(* Logix 5000 project; controller TFF vendor 1 type 14 code 107 rev 33.11; software revision 33.04; part 25 of 38 *)
(* tags used below, declared in another part *)
   Address : DINT;   // Temp Address
   Address2 : DINT;   // Temp Address
   Index : DINT;   // Index
   PCV001_PID_Settings : INT;
   TIME : DINT[2];
   AnalogOutput : AnalogOutput[25];   // Analog Output Array
   AnalogPoint : AnalogInput[50];   // Analog Input Array
   ControlLoop : ControlLoop[20];   // Control Loop Array
   ControlLoop_FeedPump : ALIAS FOR ControlLoop[1];
   ControlLoop_PCV101 : ALIAS FOR ControlLoop[3];
   ControlLoop_PCV101_5ms : ALIAS FOR ControlLoop[4];
   ControlLoop_PCV101_CV : REAL;   // Control Value
   ControlLoop_PCV101_RAMP_OUT : REAL;   // Ramp Output
   ControlLoop_PCV201 : ALIAS FOR ControlLoop[5];
   ControlLoop_PCV201_5ms : ALIAS FOR ControlLoop[6];
   ControlLoop_PCV201_RAMP_OUT : REAL;   // Ramp Output
   PCV101 : ALIAS FOR AnalogPoint[3];
   PCV101_Control : PCV_Control;   // PCV101 Control UDT
   PCV201_Control : PCV_Control;   // PCV201 Control UDT
   PumpRunStatus : DINT;   // Pumps Run Status (1 = At least one pump running , 0 = no pump running)
   SysControl : SysControl;   // General system status and command
(* Process, continued *)

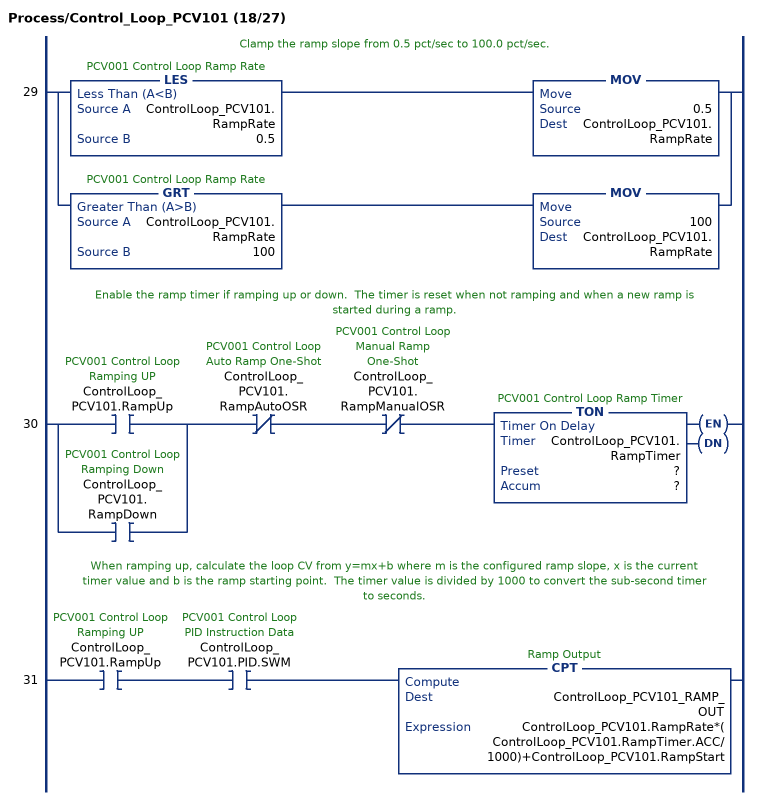
   [picture p215: Process/Control_Loop_PCV101 rungs 29-31]
   // Clamp the ramp slope from 0.5 pct/sec to 100.0 pct/sec.
   29: [LES(ControlLoop_PCV101.RampRate,0.5) MOV(0.5,ControlLoop_PCV101.RampRate) ,GRT(ControlLoop_PCV101.RampRate,100) MOV(100,ControlLoop_PCV101.RampRate) ];
   // Enable the ramp timer if ramping up or down.  The timer is reset when not ramping and when a new ramp is started during a ramp.
   30: [XIC(ControlLoop_PCV101.RampUp) ,XIC(ControlLoop_PCV101.RampDown) ]XIO(ControlLoop_PCV101.RampAutoOSR)XIO(ControlLoop_PCV101.RampManualOSR)TON(ControlLoop_PCV101.RampTimer,?,?);
   // When ramping up, calculate the loop CV from y=mx+b where m is the configured ramp slope, x is the current timer value and b is the ramp starting point.  The timer value is divided by 1000 to convert the sub-second timer to seconds.
   31: XIC(ControlLoop_PCV101.RampUp)XIC(ControlLoop_PCV101.PID.SWM)CPT(ControlLoop_PCV101_RAMP_OUT,ControlLoop_PCV101.RampRate*(ControlLoop_PCV101.RampTimer.ACC/1000)+ControlLoop_PCV101.RampStart);
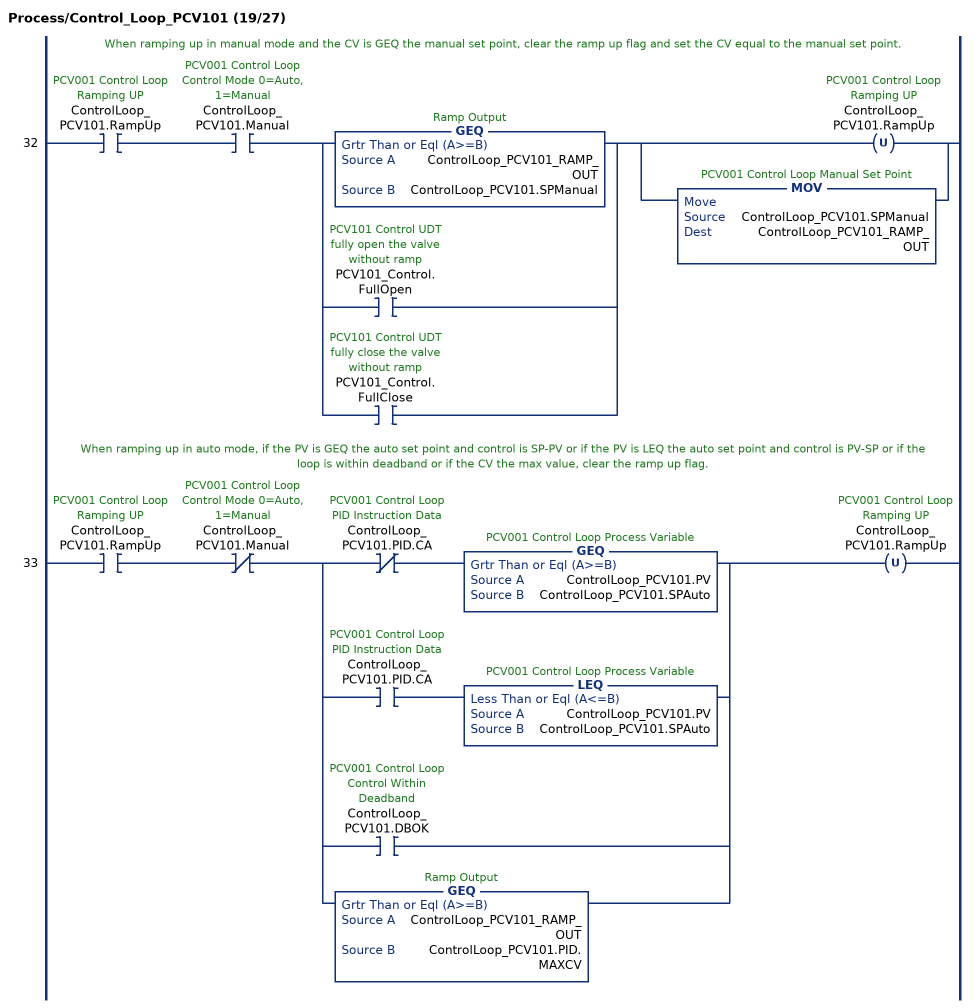
   // When ramping up in manual mode and the CV is GEQ the manual set point, clear the ramp up flag and set the CV equal to the manual set point.
   32: XIC(ControlLoop_PCV101.RampUp)XIC(ControlLoop_PCV101.Manual)[GEQ(ControlLoop_PCV101_RAMP_OUT,ControlLoop_PCV101.SPManual) ,XIC(PCV101_Control.FullOpen) ,XIC(PCV101_Control.FullClose) ][OTU(ControlLoop_PCV101.RampUp) ,MOV(ControlLoop_PCV101.SPManual,ControlLoop_PCV101_RAMP_OUT) ];
   // When ramping up in auto mode, if the PV is GEQ the auto set point and control is SP-PV or if the PV is LEQ the auto set point and control is PV-SP or if the loop is within deadband or if the CV the max value, clear the ramp up flag.
   33: XIC(ControlLoop_PCV101.RampUp)XIO(ControlLoop_PCV101.Manual)[XIO(ControlLoop_PCV101.PID.CA) GEQ(ControlLoop_PCV101.PV,ControlLoop_PCV101.SPAuto) ,XIC(ControlLoop_PCV101.PID.CA) LEQ(ControlLoop_PCV101.PV,ControlLoop_PCV101.SPAuto) ,XIC(ControlLoop_PCV101.DBOK) ,GEQ(ControlLoop_PCV101_RAMP_OUT,ControlLoop_PCV101.PID.MAXCV) ]OTU(ControlLoop_PCV101.RampUp);
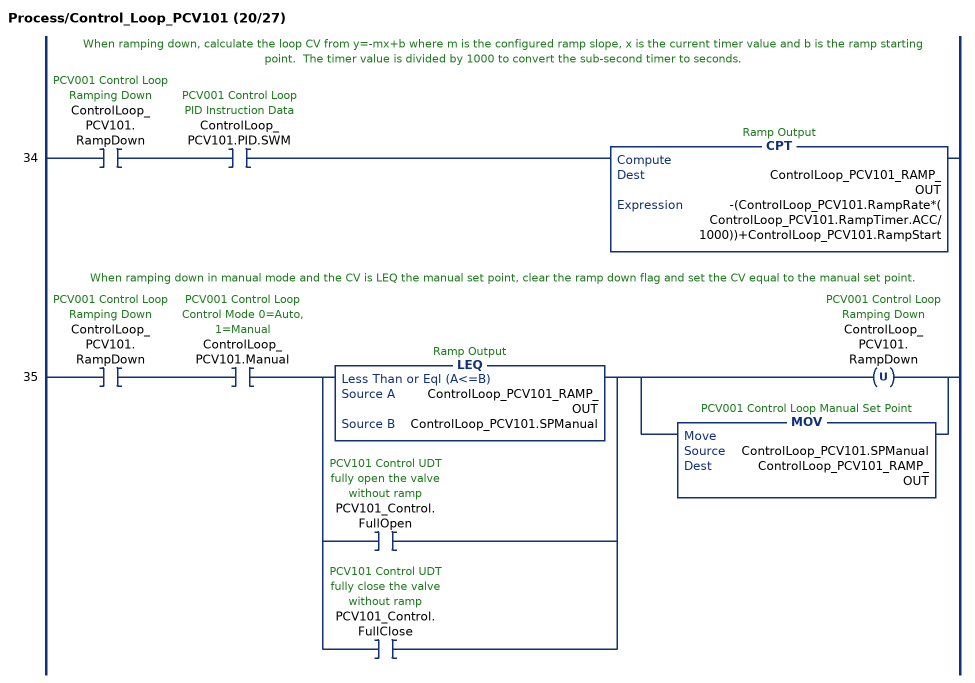
   // When ramping down, calculate the loop CV from y=-mx+b where m is the configured ramp slope, x is the current timer value and b is the ramp starting point.  The timer value is divided by 1000 to convert the sub-second timer to seconds.
   34: XIC(ControlLoop_PCV101.RampDown)XIC(ControlLoop_PCV101.PID.SWM)CPT(ControlLoop_PCV101_RAMP_OUT,-(ControlLoop_PCV101.RampRate*(ControlLoop_PCV101.RampTimer.ACC/1000))+ControlLoop_PCV101.RampStart);
   // When ramping down in manual mode and the CV is LEQ the manual set point, clear the ramp down flag and set the CV equal to the manual set point.
   35: XIC(ControlLoop_PCV101.RampDown)XIC(ControlLoop_PCV101.Manual)[LEQ(ControlLoop_PCV101_RAMP_OUT,ControlLoop_PCV101.SPManual) ,XIC(PCV101_Control.FullOpen) ,XIC(PCV101_Control.FullClose) ][OTU(ControlLoop_PCV101.RampDown) ,MOV(ControlLoop_PCV101.SPManual,ControlLoop_PCV101_RAMP_OUT) ];
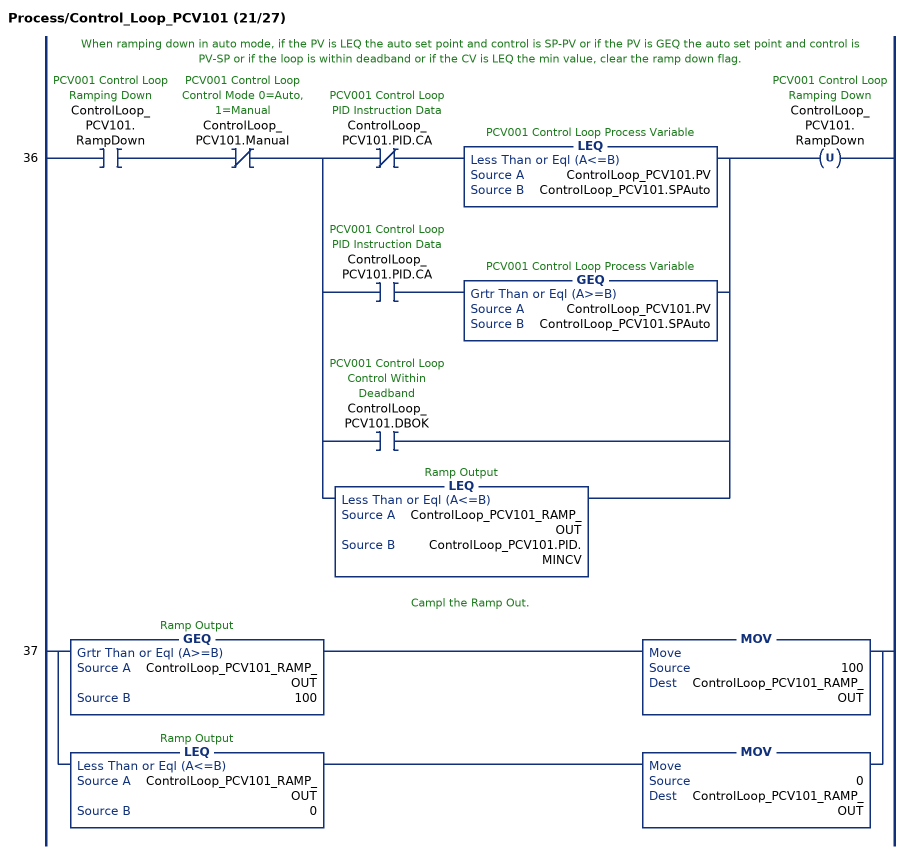
   // When ramping down in auto mode, if the PV is LEQ the auto set point and control is SP-PV or if the PV is GEQ the auto set point and control is PV-SP or if the loop is within deadband or if the CV is LEQ the min value, clear the ramp down flag.
   36: XIC(ControlLoop_PCV101.RampDown)XIO(ControlLoop_PCV101.Manual)[XIO(ControlLoop_PCV101.PID.CA) LEQ(ControlLoop_PCV101.PV,ControlLoop_PCV101.SPAuto) ,XIC(ControlLoop_PCV101.PID.CA) GEQ(ControlLoop_PCV101.PV,ControlLoop_PCV101.SPAuto) ,XIC(ControlLoop_PCV101.DBOK) ,LEQ(ControlLoop_PCV101_RAMP_OUT,ControlLoop_PCV101.PID.MINCV) ]OTU(ControlLoop_PCV101.RampDown);
   // Campl the Ramp Out.
   37: [GEQ(ControlLoop_PCV101_RAMP_OUT,100) MOV(100,ControlLoop_PCV101_RAMP_OUT) ,LEQ(ControlLoop_PCV101_RAMP_OUT,0) MOV(0,ControlLoop_PCV101_RAMP_OUT) ];
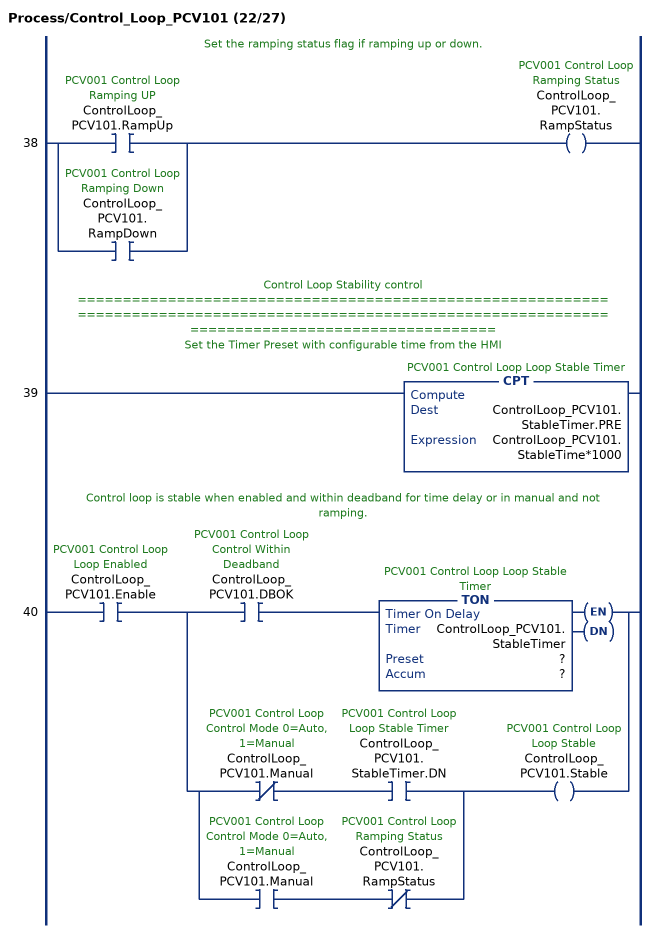
   // Set the ramping status flag if ramping up or down.
   38: [XIC(ControlLoop_PCV101.RampUp) ,XIC(ControlLoop_PCV101.RampDown) ]OTE(ControlLoop_PCV101.RampStatus);
   // Control Loop Stability control
   // ========================================================================================================================================================
   // Set the Timer Preset with configurable time from the HMI
   39: CPT(ControlLoop_PCV101.StableTimer.PRE,ControlLoop_PCV101.StableTime*1000);
   // Control loop is stable when enabled and within deadband for time delay or in manual and not ramping.
   40: XIC(ControlLoop_PCV101.Enable)[XIC(ControlLoop_PCV101.DBOK) TON(ControlLoop_PCV101.StableTimer,?,?) ,[XIO(ControlLoop_PCV101.Manual) XIC(ControlLoop_PCV101.StableTimer.DN) ,XIC(ControlLoop_PCV101.Manual) XIO(ControlLoop_PCV101.RampStatus) ] OTE(ControlLoop_PCV101.Stable) ];
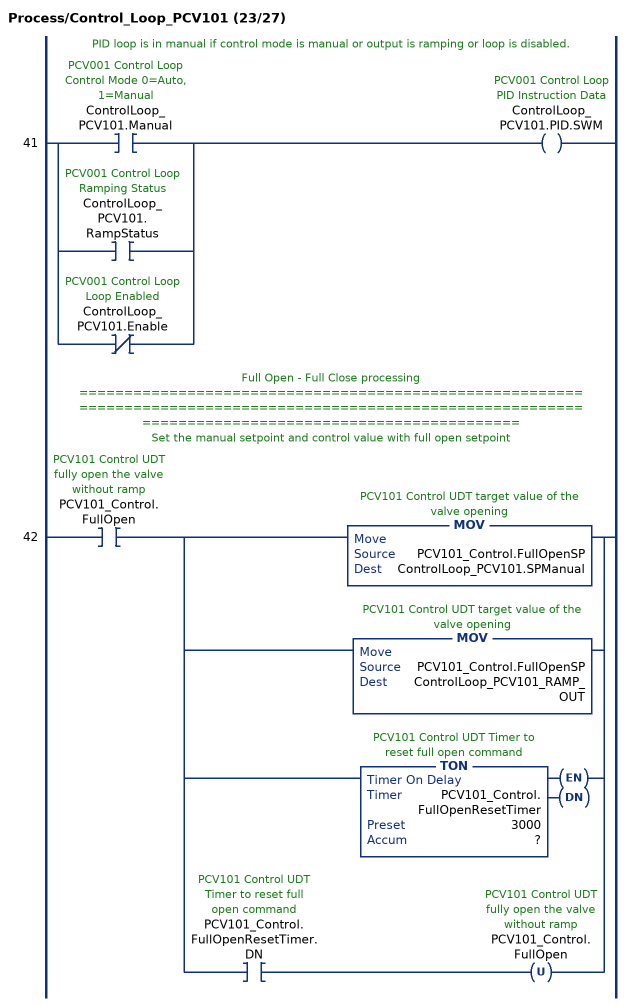
   // PID loop is in manual if control mode is manual or output is ramping or loop is disabled.
   41: [XIC(ControlLoop_PCV101.Manual) ,XIC(ControlLoop_PCV101.RampStatus) ,XIO(ControlLoop_PCV101.Enable) ]OTE(ControlLoop_PCV101.PID.SWM);
   // Full Open - Full Close processing
   // ==========================================================================================================================================================
   // Set the manual setpoint and control value with full open setpoint
   42: XIC(PCV101_Control.FullOpen)[MOV(PCV101_Control.FullOpenSP,ControlLoop_PCV101.SPManual) ,MOV(PCV101_Control.FullOpenSP,ControlLoop_PCV101_RAMP_OUT) ,TON(PCV101_Control.FullOpenResetTimer,?,?) ,XIC(PCV101_Control.FullOpenResetTimer.DN) OTU(PCV101_Control.FullOpen) ];
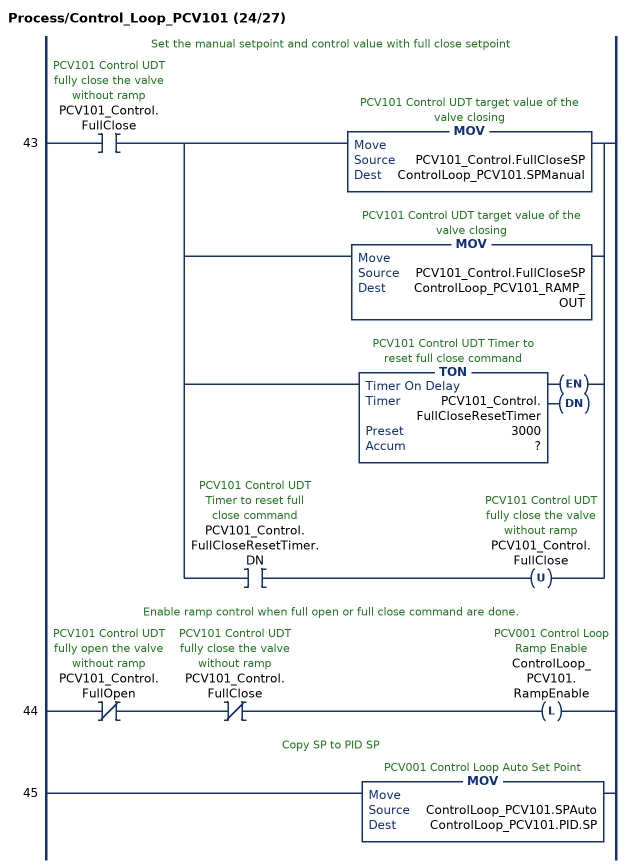
   // Set the manual setpoint and control value with full close setpoint
   43: XIC(PCV101_Control.FullClose)[MOV(PCV101_Control.FullCloseSP,ControlLoop_PCV101.SPManual) ,MOV(PCV101_Control.FullCloseSP,ControlLoop_PCV101_RAMP_OUT) ,TON(PCV101_Control.FullCloseResetTimer,?,?) ,XIC(PCV101_Control.FullCloseResetTimer.DN) OTU(PCV101_Control.FullClose) ];
   // Enable ramp control when full open or full close command are done.
   44: XIO(PCV101_Control.FullOpen)XIO(PCV101_Control.FullClose)OTL(ControlLoop_PCV101.RampEnable);
   // Copy SP to PID SP
   45: MOV(ControlLoop_PCV101.SPAuto,ControlLoop_PCV101.PID.SP);
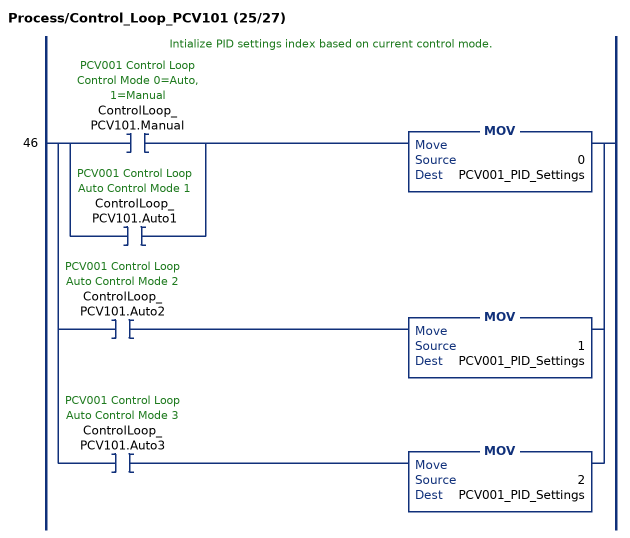
   // Intialize PID settings index based on current control mode.
   46: [[XIC(ControlLoop_PCV101.Manual) ,XIC(ControlLoop_PCV101.Auto1) ] MOV(0,PCV001_PID_Settings) ,XIC(ControlLoop_PCV101.Auto2) MOV(1,PCV001_PID_Settings) ,XIC(ControlLoop_PCV101.Auto3) MOV(2,PCV001_PID_Settings) ];
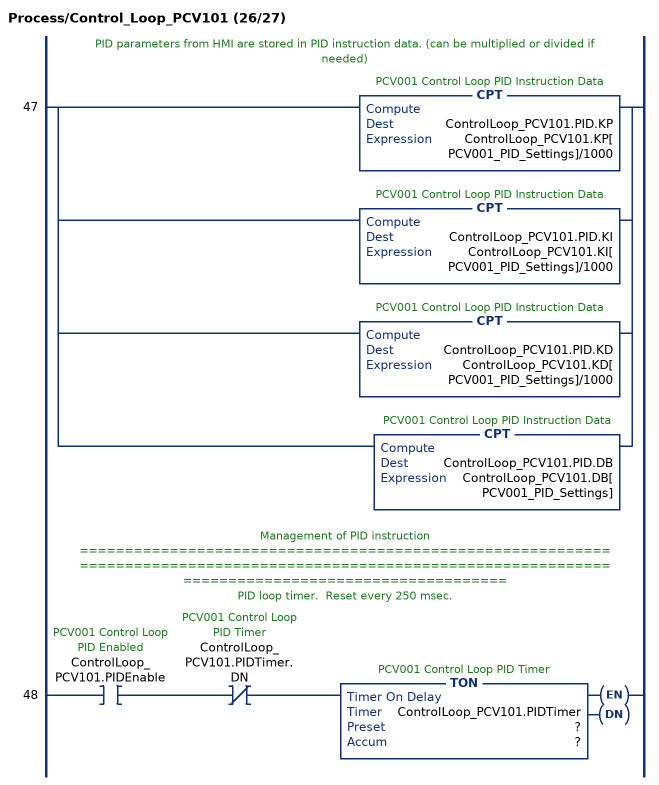
   // PID parameters from HMI are stored in PID instruction data. (can be multiplied or divided if needed)
   47: [CPT(ControlLoop_PCV101.PID.KP,ControlLoop_PCV101.KP[PCV001_PID_Settings]/1000) ,CPT(ControlLoop_PCV101.PID.KI,ControlLoop_PCV101.KI[PCV001_PID_Settings]/1000) ,CPT(ControlLoop_PCV101.PID.KD,ControlLoop_PCV101.KD[PCV001_PID_Settings]/1000) ,CPT(ControlLoop_PCV101.PID.DB,ControlLoop_PCV101.DB[PCV001_PID_Settings]) ];
   // Management of PID instruction
   // ==========================================================================================================================================================
   // PID loop timer.  Reset every 250 msec.
   48: XIC(ControlLoop_PCV101.PIDEnable)XIO(ControlLoop_PCV101.PIDTimer.DN)TON(ControlLoop_PCV101.PIDTimer,?,?);
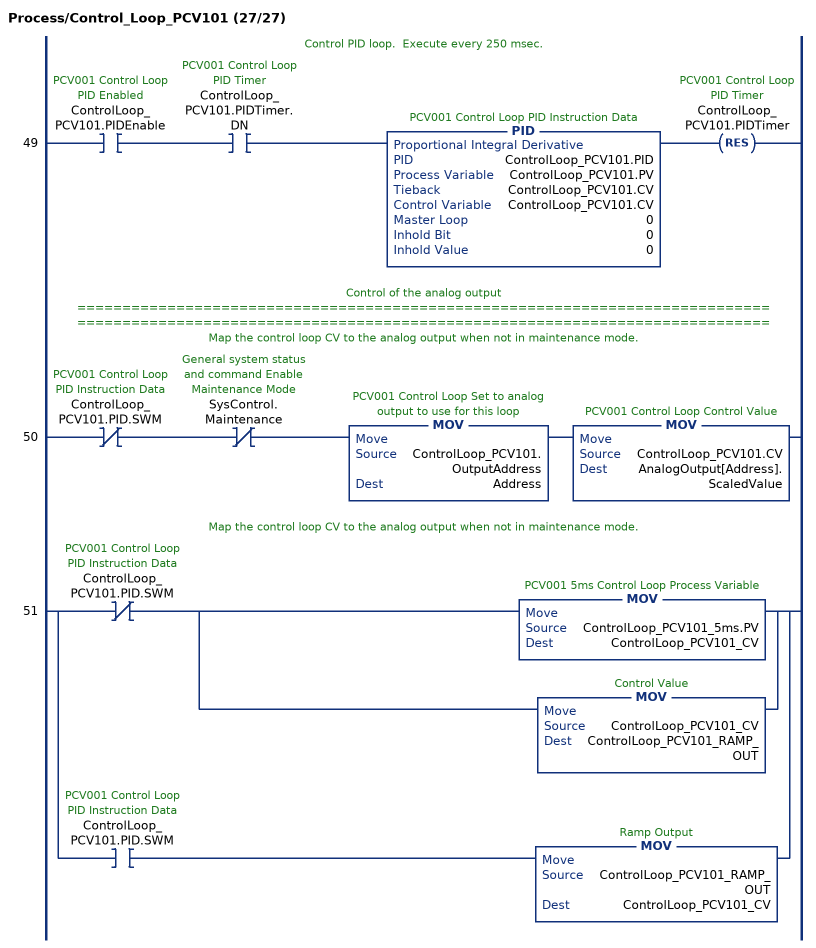
   // Control PID loop.  Execute every 250 msec.
   49: XIC(ControlLoop_PCV101.PIDEnable)XIC(ControlLoop_PCV101.PIDTimer.DN)PID(ControlLoop_PCV101.PID,ControlLoop_PCV101.PV,ControlLoop_PCV101.CV,ControlLoop_PCV101.CV,0,0,0)RES(ControlLoop_PCV101.PIDTimer);
   // Control of the analog output
   // ==========================================================================================================================================================
   // Map the control loop CV to the analog output when not in maintenance mode.
   50: XIO(ControlLoop_PCV101.PID.SWM)XIO(SysControl.Maintenance)MOV(ControlLoop_PCV101.OutputAddress,Address)MOV(ControlLoop_PCV101.CV,AnalogOutput[Address].ScaledValue);
   // Map the control loop CV to the analog output when not in maintenance mode.
   51: [XIO(ControlLoop_PCV101.PID.SWM) [MOV(ControlLoop_PCV101_5ms.PV,ControlLoop_PCV101_CV) ,MOV(ControlLoop_PCV101_CV,ControlLoop_PCV101_RAMP_OUT) ] ,XIC(ControlLoop_PCV101.PID.SWM) MOV(ControlLoop_PCV101_RAMP_OUT,ControlLoop_PCV101_CV) ];
END_ROUTINE

ROUTINE Control_Loop_PCV201   (* ladder *)
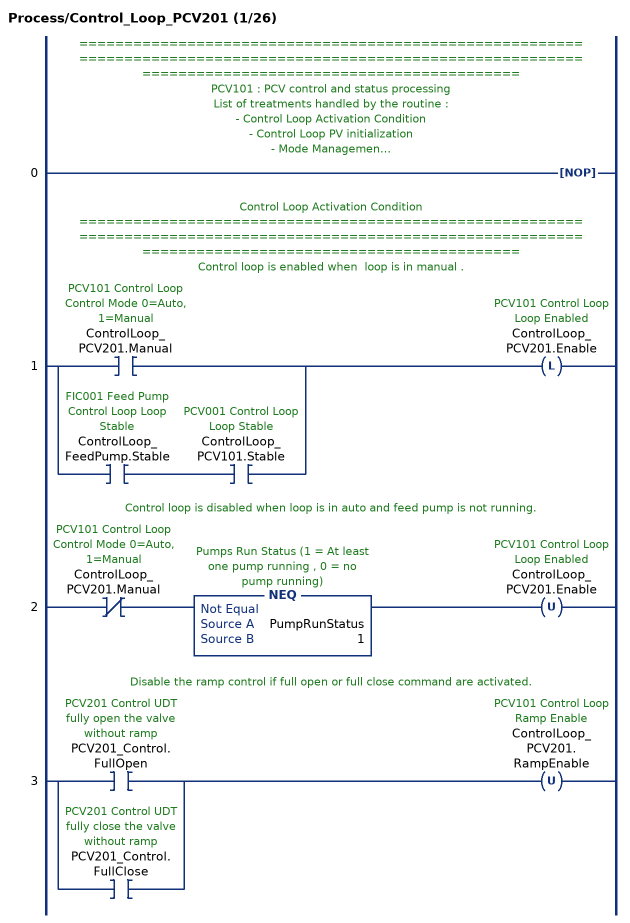
   // ==========================================================================================================================================================
   //                                                  PCV101 : PCV control and status processing
   //                                                     List of treatments handled by the routine :
   //                                                          - Control Loop Activation Condition
   //                                                  - Control Loop PV initialization
   //                                                - Mode Management
   //                                                        - Control Loop Setpoint management
   //                                                        - Control Loop deadband calculation
   //                                                          - Management of ramping control
   //                                                          - Control Loop Stability control
   //                                                          - Full Open - Full Close processing
   //                                                          - Management of PID instruction
   //                                                          - Control of the analog output
   //                                                     -----------------------------------------------------------------------------------------------------------------------------------------------------
   //                                                     History
   // 		2019-DEC-24 - Merck - Q. Spindler - Initial version for Candidate Release 1.00.00.00.a
   // 		2020-SEP-09 - Merck - Q. Spindler - Modifications for Candidate Release 1.00.00.00.d
   // 					- Add ControlLoop Enable and not manual condition for DBOK status
   // 		2021-APR-16 - Merck - Q. Spindler - Modifications for Candidate Release 1.00.00.00.e
   //                                        - Add Initialize address if no mode selected.
   // ==========================================================================================================================================================
   0: NOP();
   // Control Loop Activation Condition
   // ==========================================================================================================================================================
   // Control loop is enabled when  loop is in manual .
   1: [XIC(ControlLoop_PCV201.Manual) ,XIC(ControlLoop_FeedPump.Stable) XIC(ControlLoop_PCV101.Stable) ]OTL(ControlLoop_PCV201.Enable);
   // Control loop is disabled when loop is in auto and feed pump is not running.
   2: XIO(ControlLoop_PCV201.Manual)NEQ(PumpRunStatus,1)OTU(ControlLoop_PCV201.Enable);
   // Disable the ramp control if full open or full close command are activated.
   3: [XIC(PCV201_Control.FullOpen) ,XIC(PCV201_Control.FullClose) ]OTU(ControlLoop_PCV201.RampEnable);
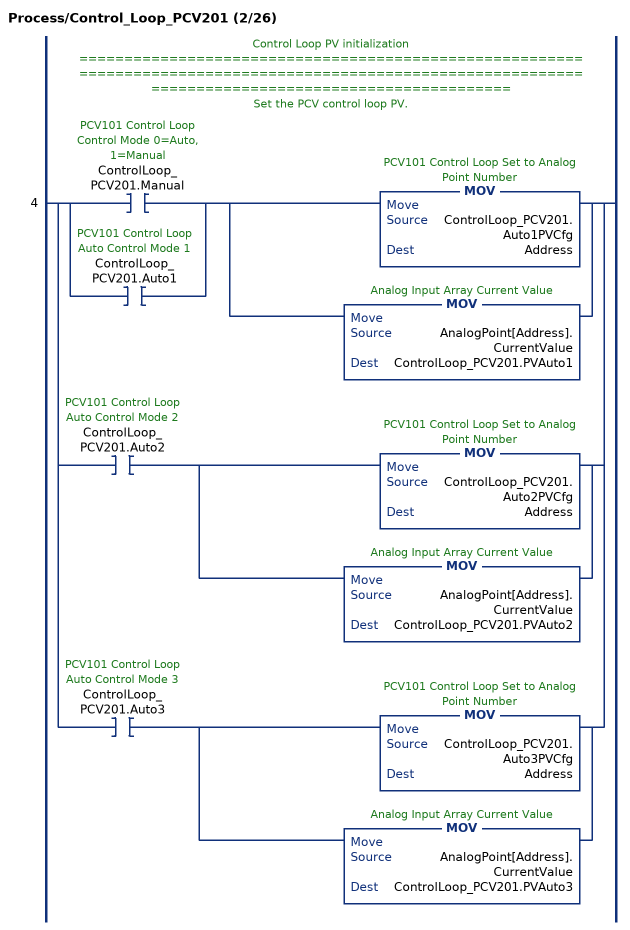
   // Control Loop PV initialization
   // ========================================================================================================================================================
   // Set the PCV control loop PV.
   4: [[[XIC(ControlLoop_PCV201.Manual) ,XIC(ControlLoop_PCV201.Auto1) ] [MOV(ControlLoop_PCV201.Auto1PVCfg,Address) ,MOV(AnalogPoint[Address].CurrentValue,ControlLoop_PCV201.PVAuto1) ] ,XIC(ControlLoop_PCV201.Auto2) [MOV(ControlLoop_PCV201.Auto2PVCfg,Address) ,MOV(AnalogPoint[Address].CurrentValue,ControlLoop_PCV201.PVAuto2) ] ] ,XIC(ControlLoop_PCV201.Auto3) [MOV(ControlLoop_PCV201.Auto3PVCfg,Address) ,MOV(AnalogPoint[Address].CurrentValue,ControlLoop_PCV201.PVAuto3) ] ];
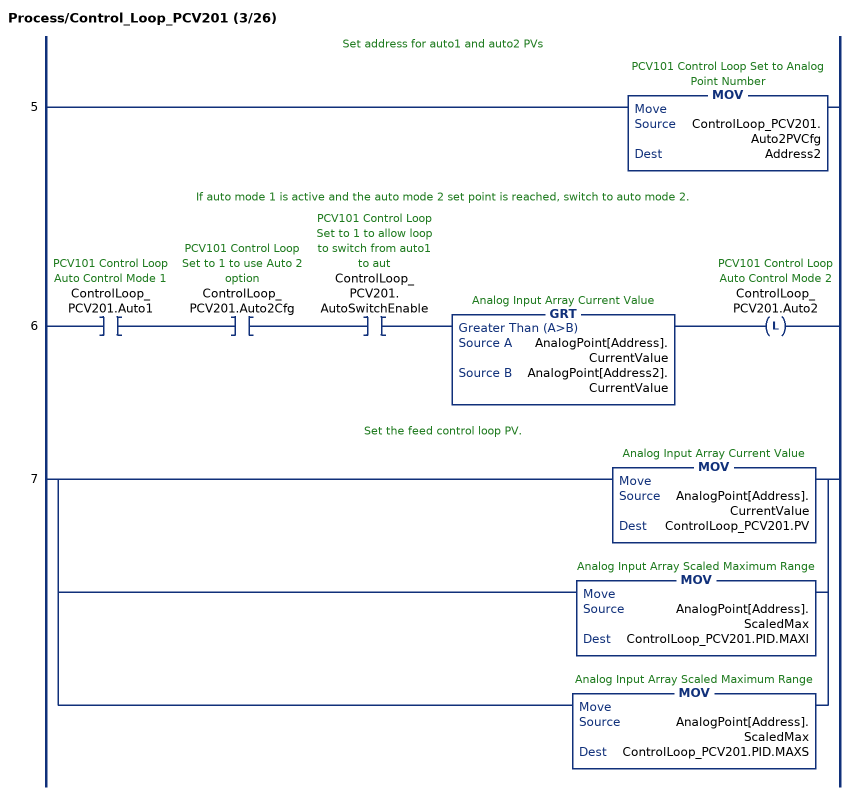
   // Set address for auto1 and auto2 PVs
   5: MOV(ControlLoop_PCV201.Auto2PVCfg,Address2);
   // If auto mode 1 is active and the auto mode 2 set point is reached, switch to auto mode 2.
   6: XIC(ControlLoop_PCV201.Auto1)XIC(ControlLoop_PCV201.Auto2Cfg)XIC(ControlLoop_PCV201.AutoSwitchEnable)GRT(AnalogPoint[Address].CurrentValue,AnalogPoint[Address2].CurrentValue)OTL(ControlLoop_PCV201.Auto2);
   // Set the feed control loop PV.
   7: [MOV(AnalogPoint[Address].CurrentValue,ControlLoop_PCV201.PV) ,MOV(AnalogPoint[Address].ScaledMax,ControlLoop_PCV201.PID.MAXI) ,MOV(AnalogPoint[Address].ScaledMax,ControlLoop_PCV201.PID.MAXS) ];
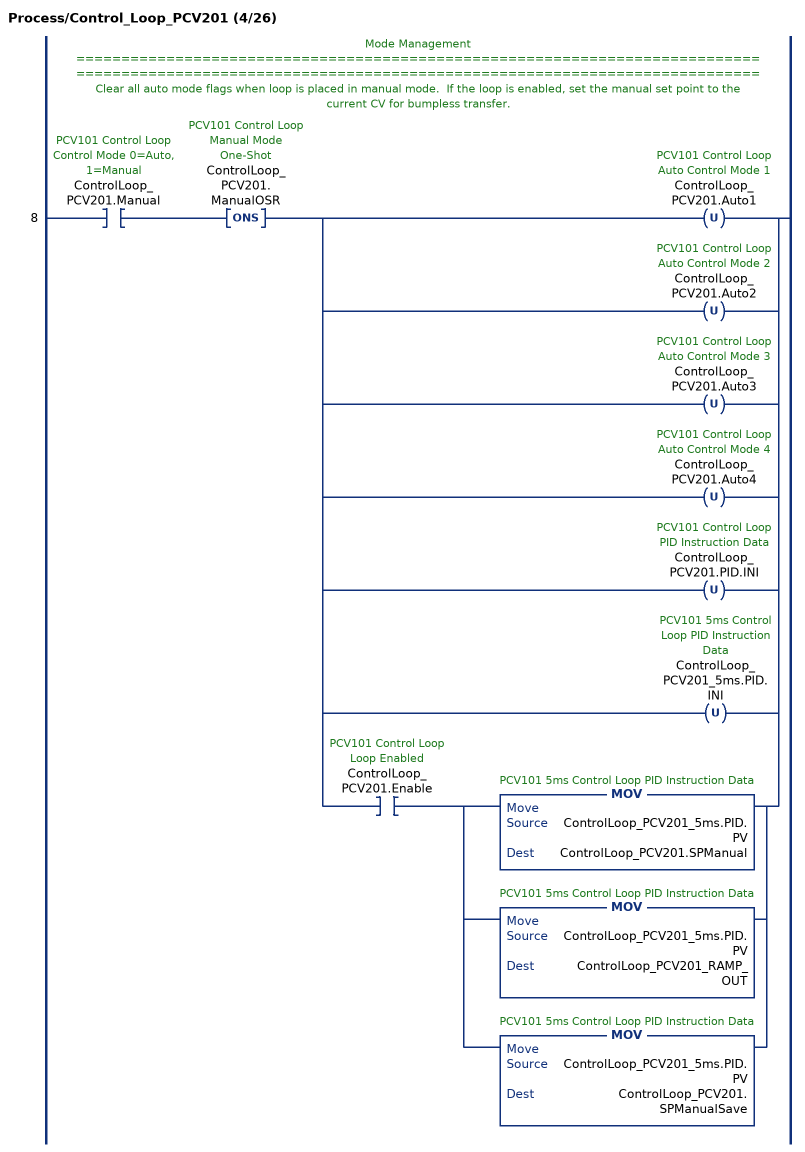
   // Mode Management
   // ========================================================================================================================================================
   // Clear all auto mode flags when loop is placed in manual mode.  If the loop is enabled, set the manual set point to the current CV for bumpless transfer.
   8: XIC(ControlLoop_PCV201.Manual)ONS(ControlLoop_PCV201.ManualOSR)[OTU(ControlLoop_PCV201.Auto1) ,OTU(ControlLoop_PCV201.Auto2) ,OTU(ControlLoop_PCV201.Auto3) ,OTU(ControlLoop_PCV201.Auto4) ,OTU(ControlLoop_PCV201.PID.INI) ,OTU(ControlLoop_PCV201_5ms.PID.INI) ,XIC(ControlLoop_PCV201.Enable) [MOV(ControlLoop_PCV201_5ms.PID.PV,ControlLoop_PCV201.SPManual) ,MOV(ControlLoop_PCV201_5ms.PID.PV,ControlLoop_PCV201_RAMP_OUT) ,MOV(ControlLoop_PCV201_5ms.PID.PV,ControlLoop_PCV201.SPManualSave) ] ];
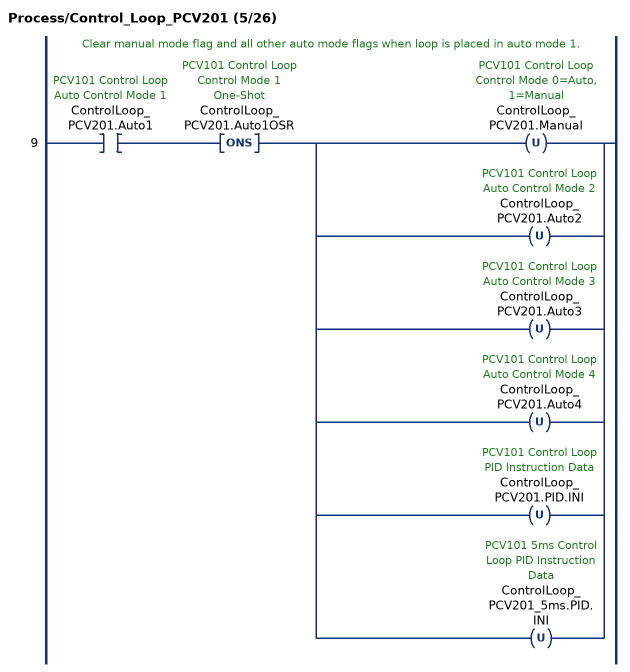
   // Clear manual mode flag and all other auto mode flags when loop is placed in auto mode 1.
   9: XIC(ControlLoop_PCV201.Auto1)ONS(ControlLoop_PCV201.Auto1OSR)[OTU(ControlLoop_PCV201.Manual) ,OTU(ControlLoop_PCV201.Auto2) ,OTU(ControlLoop_PCV201.Auto3) ,OTU(ControlLoop_PCV201.Auto4) ,OTU(ControlLoop_PCV201.PID.INI) ,OTU(ControlLoop_PCV201_5ms.PID.INI) ];
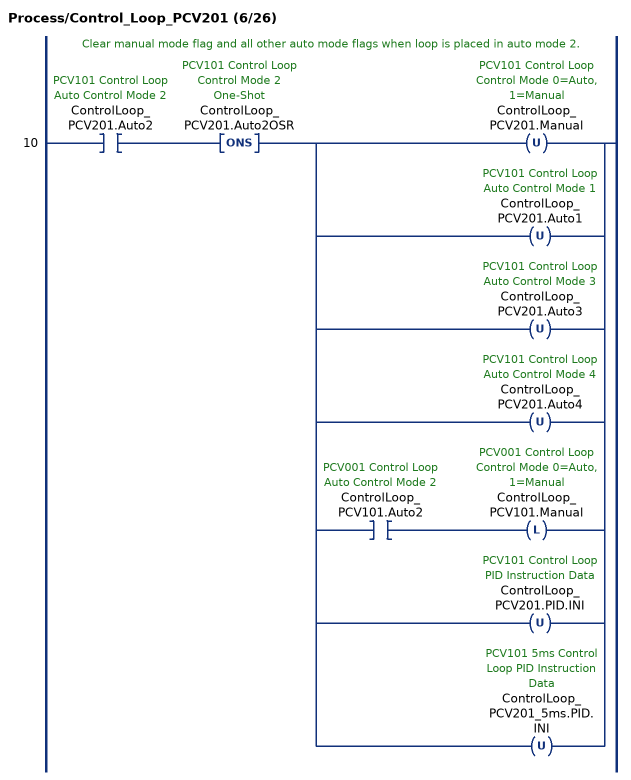
   // Clear manual mode flag and all other auto mode flags when loop is placed in auto mode 2.
   10: XIC(ControlLoop_PCV201.Auto2)ONS(ControlLoop_PCV201.Auto2OSR)[OTU(ControlLoop_PCV201.Manual) ,OTU(ControlLoop_PCV201.Auto1) ,OTU(ControlLoop_PCV201.Auto3) ,OTU(ControlLoop_PCV201.Auto4) ,XIC(ControlLoop_PCV101.Auto2) OTL(ControlLoop_PCV101.Manual) ,OTU(ControlLoop_PCV201.PID.INI) ,OTU(ControlLoop_PCV201_5ms.PID.INI) ];
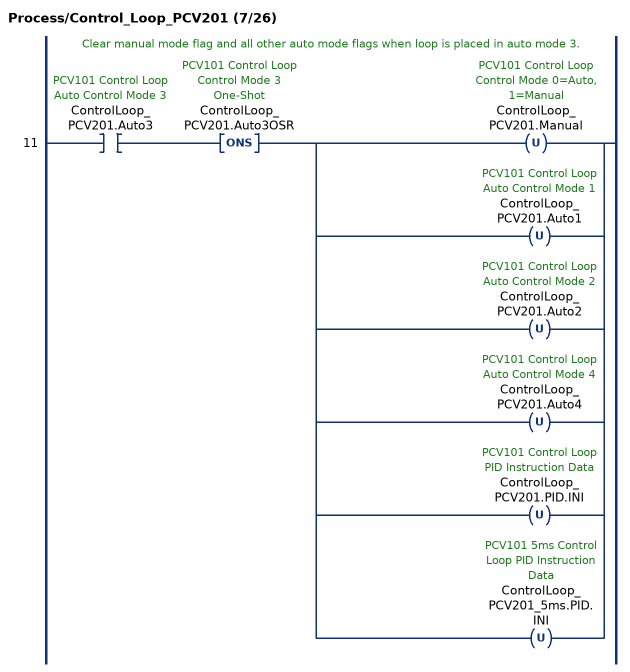
   // Clear manual mode flag and all other auto mode flags when loop is placed in auto mode 3.
   11: XIC(ControlLoop_PCV201.Auto3)ONS(ControlLoop_PCV201.Auto3OSR)[OTU(ControlLoop_PCV201.Manual) ,OTU(ControlLoop_PCV201.Auto1) ,OTU(ControlLoop_PCV201.Auto2) ,OTU(ControlLoop_PCV201.Auto4) ,OTU(ControlLoop_PCV201.PID.INI) ,OTU(ControlLoop_PCV201_5ms.PID.INI) ];
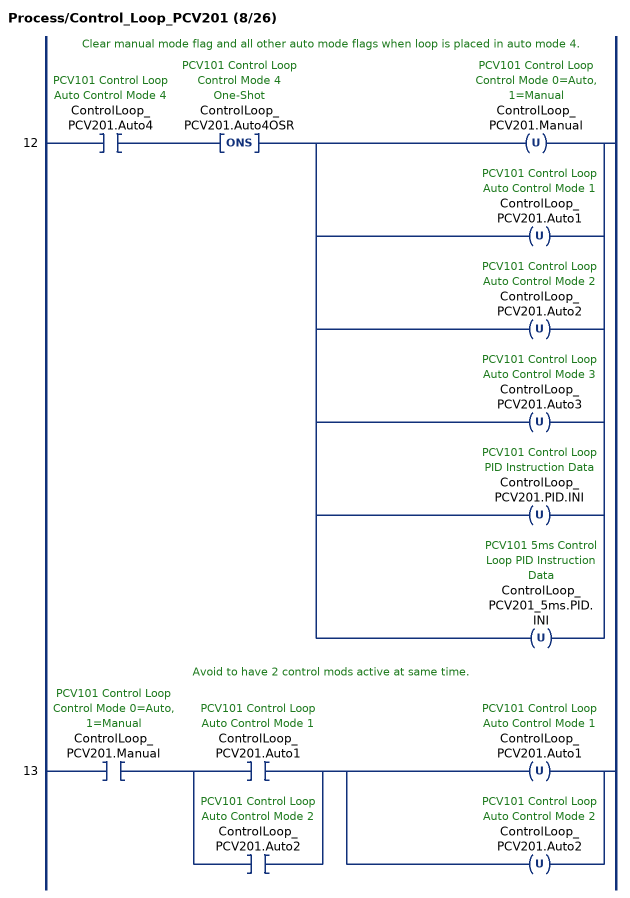
   // Clear manual mode flag and all other auto mode flags when loop is placed in auto mode 4.
   12: XIC(ControlLoop_PCV201.Auto4)ONS(ControlLoop_PCV201.Auto4OSR)[OTU(ControlLoop_PCV201.Manual) ,OTU(ControlLoop_PCV201.Auto1) ,OTU(ControlLoop_PCV201.Auto2) ,OTU(ControlLoop_PCV201.Auto3) ,OTU(ControlLoop_PCV201.PID.INI) ,OTU(ControlLoop_PCV201_5ms.PID.INI) ];
   // Avoid to have 2 control mods active at same time.
   13: XIC(ControlLoop_PCV201.Manual)[XIC(ControlLoop_PCV201.Auto1) ,XIC(ControlLoop_PCV201.Auto2) ][OTU(ControlLoop_PCV201.Auto1) ,OTU(ControlLoop_PCV201.Auto2) ];
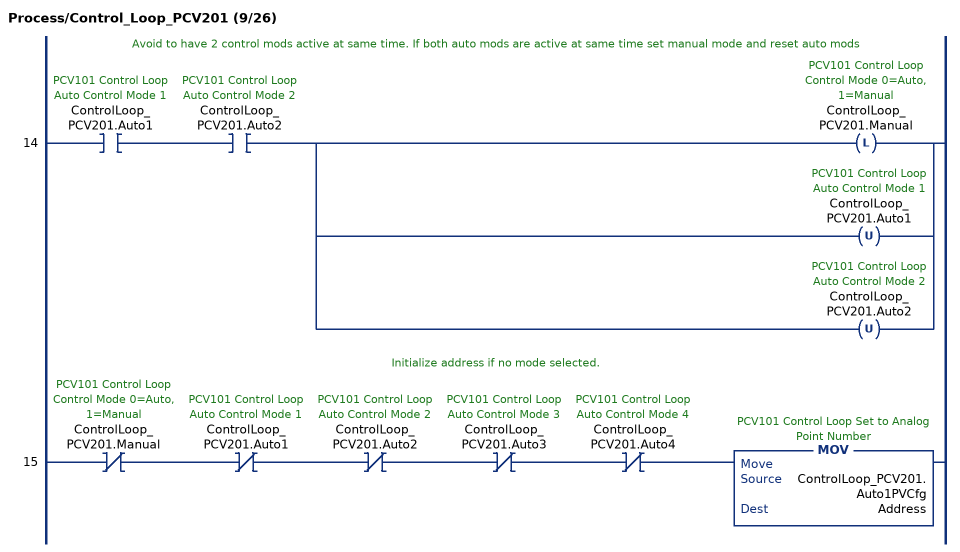
   // Avoid to have 2 control mods active at same time. If both auto mods are active at same time set manual mode and reset auto mods
   14: XIC(ControlLoop_PCV201.Auto1)XIC(ControlLoop_PCV201.Auto2)[OTL(ControlLoop_PCV201.Manual) ,OTU(ControlLoop_PCV201.Auto1) ,OTU(ControlLoop_PCV201.Auto2) ];
   // Initialize address if no mode selected.
   15: XIO(ControlLoop_PCV201.Manual)XIO(ControlLoop_PCV201.Auto1)XIO(ControlLoop_PCV201.Auto2)XIO(ControlLoop_PCV201.Auto3)XIO(ControlLoop_PCV201.Auto4)MOV(ControlLoop_PCV201.Auto1PVCfg,Address);
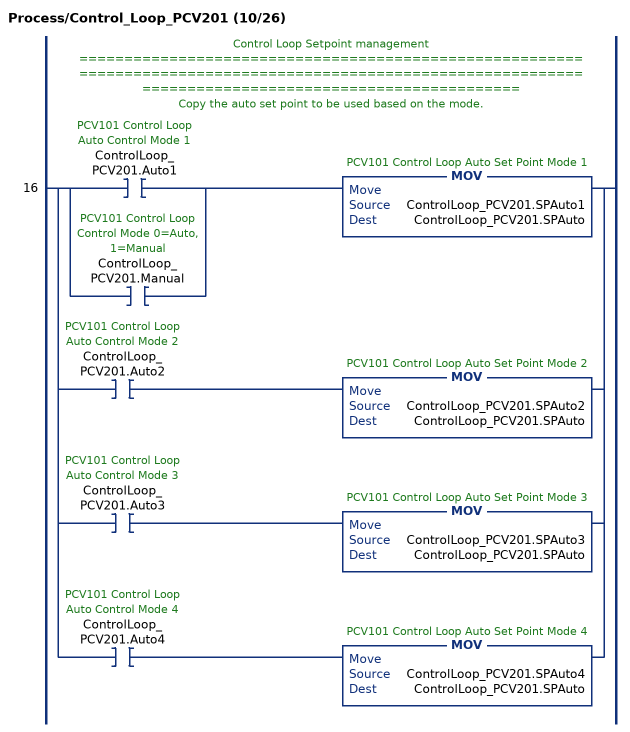
   // Control Loop Setpoint management
   // ==========================================================================================================================================================
   // Copy the auto set point to be used based on the mode.
   16: [[XIC(ControlLoop_PCV201.Auto1) ,XIC(ControlLoop_PCV201.Manual) ] MOV(ControlLoop_PCV201.SPAuto1,ControlLoop_PCV201.SPAuto) ,XIC(ControlLoop_PCV201.Auto2) MOV(ControlLoop_PCV201.SPAuto2,ControlLoop_PCV201.SPAuto) ,XIC(ControlLoop_PCV201.Auto3) MOV(ControlLoop_PCV201.SPAuto3,ControlLoop_PCV201.SPAuto) ,XIC(ControlLoop_PCV201.Auto4) MOV(ControlLoop_PCV201.SPAuto4,ControlLoop_PCV201.SPAuto) ];
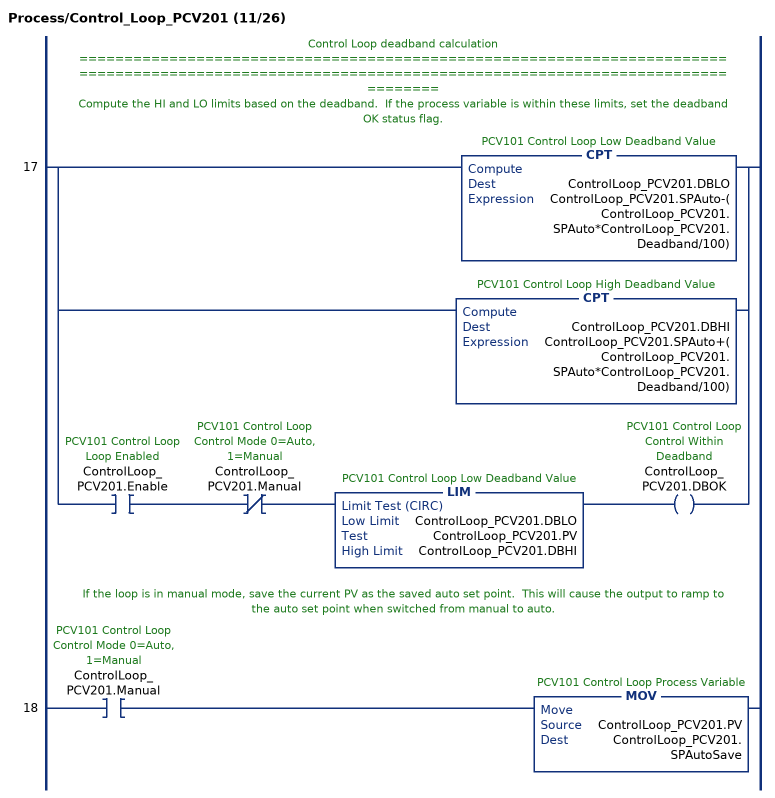
   // Control Loop deadband calculation
   // ========================================================================================================================================================
   // Compute the HI and LO limits based on the deadband.  If the process variable is within these limits, set the deadband OK status flag.
   17: [CPT(ControlLoop_PCV201.DBLO,ControlLoop_PCV201.SPAuto-(ControlLoop_PCV201.SPAuto*ControlLoop_PCV201.Deadband/100)) ,CPT(ControlLoop_PCV201.DBHI,ControlLoop_PCV201.SPAuto+(ControlLoop_PCV201.SPAuto*ControlLoop_PCV201.Deadband/100)) ,XIC(ControlLoop_PCV201.Enable) XIO(ControlLoop_PCV201.Manual) LIM(ControlLoop_PCV201.DBLO,ControlLoop_PCV201.PV,ControlLoop_PCV201.DBHI) OTE(ControlLoop_PCV201.DBOK) ];
   // If the loop is in manual mode, save the current PV as the saved auto set point.  This will cause the output to ramp to the auto set point when switched from manual to auto.
   18: XIC(ControlLoop_PCV201.Manual)MOV(ControlLoop_PCV201.PV,ControlLoop_PCV201.SPAutoSave);
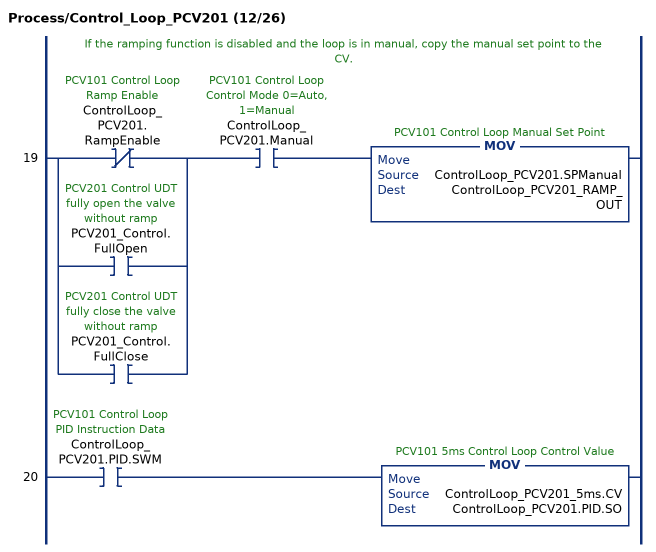
   // If the ramping function is disabled and the loop is in manual, copy the manual set point to the CV.
   19: [XIO(ControlLoop_PCV201.RampEnable) ,XIC(PCV201_Control.FullOpen) ,XIC(PCV201_Control.FullClose) ]XIC(ControlLoop_PCV201.Manual)MOV(ControlLoop_PCV201.SPManual,ControlLoop_PCV201_RAMP_OUT);
   20: XIC(ControlLoop_PCV201.PID.SWM)MOV(ControlLoop_PCV201_5ms.CV,ControlLoop_PCV201.PID.SO);
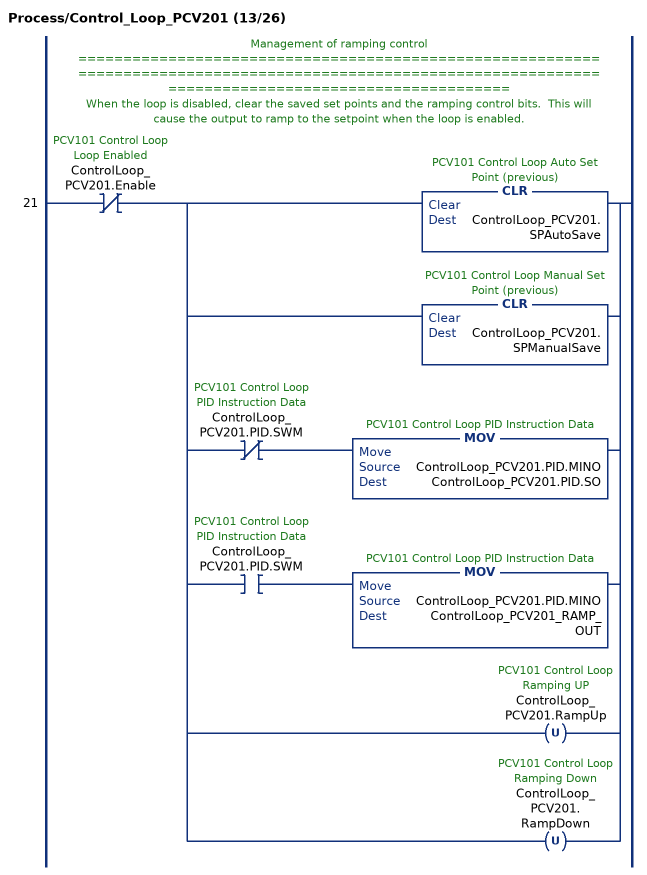
   // Management of ramping control
   // ==========================================================================================================================================================
   // When the loop is disabled, clear the saved set points and the ramping control bits.  This will cause the output to ramp to the setpoint when the loop is enabled.
   21: XIO(ControlLoop_PCV201.Enable)[CLR(ControlLoop_PCV201.SPAutoSave) ,CLR(ControlLoop_PCV201.SPManualSave) ,XIO(ControlLoop_PCV201.PID.SWM) MOV(ControlLoop_PCV201.PID.MINO,ControlLoop_PCV201.PID.SO) ,XIC(ControlLoop_PCV201.PID.SWM) MOV(ControlLoop_PCV201.PID.MINO,ControlLoop_PCV201_RAMP_OUT) ,OTU(ControlLoop_PCV201.RampUp) ,OTU(ControlLoop_PCV201.RampDown) ];
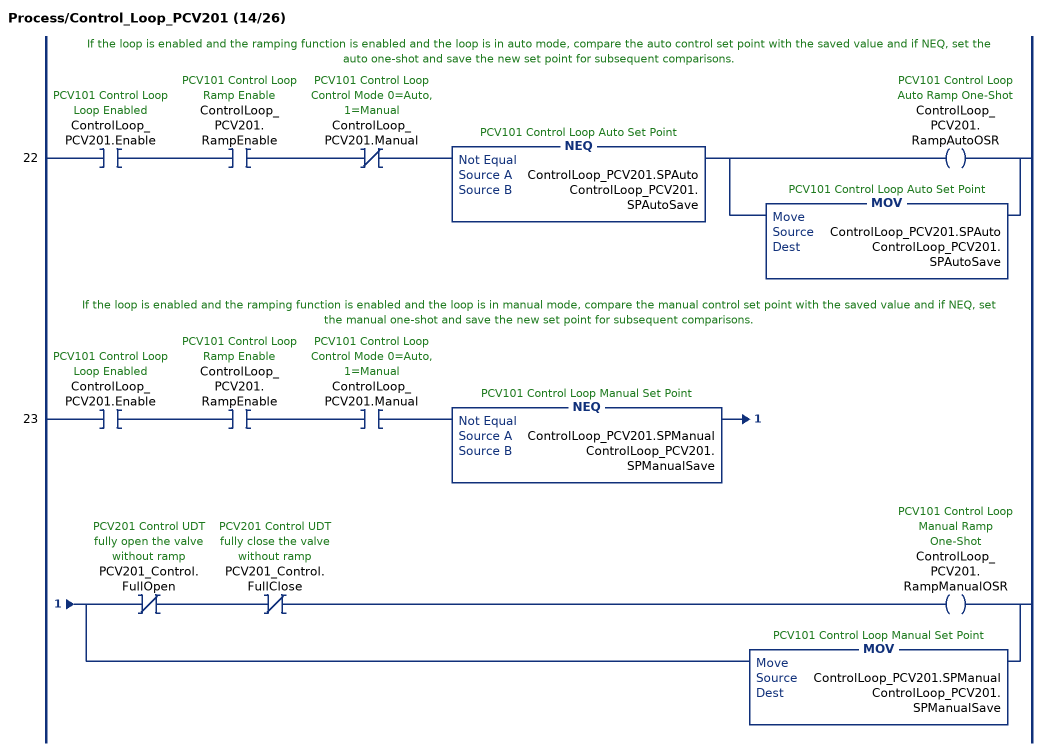
   // If the loop is enabled and the ramping function is enabled and the loop is in auto mode, compare the auto control set point with the saved value and if NEQ, set the auto one-shot and save the new set point for subsequent comparisons.
   22: XIC(ControlLoop_PCV201.Enable)XIC(ControlLoop_PCV201.RampEnable)XIO(ControlLoop_PCV201.Manual)NEQ(ControlLoop_PCV201.SPAuto,ControlLoop_PCV201.SPAutoSave)[OTE(ControlLoop_PCV201.RampAutoOSR) ,MOV(ControlLoop_PCV201.SPAuto,ControlLoop_PCV201.SPAutoSave) ];
   // If the loop is enabled and the ramping function is enabled and the loop is in manual mode, compare the manual control set point with the saved value and if NEQ, set the manual one-shot and save the new set point for subsequent comparisons.
   23: XIC(ControlLoop_PCV201.Enable)XIC(ControlLoop_PCV201.RampEnable)XIC(ControlLoop_PCV201.Manual)NEQ(ControlLoop_PCV201.SPManual,ControlLoop_PCV201.SPManualSave)[XIO(PCV201_Control.FullOpen) XIO(PCV201_Control.FullClose) OTE(ControlLoop_PCV201.RampManualOSR) ,MOV(ControlLoop_PCV201.SPManual,ControlLoop_PCV201.SPManualSave) ];
